PROGRAM main
  VAR
    B1 AT %IX0.0  : BOOL; (* sensor de piezas *)
    S1 AT %IX0.1  : BOOL; (* RESET *)
    KM1 AT %QX0.0 : BOOL; (* motor de la cinta *)
    H1 AT %QX0.1  : BOOL; (* caja llena *)
    PIEZAS        : CTU;
    LLENA         : BOOL;
    CUENTA        : INT; (* piezas en la caja *)
  END_VAR

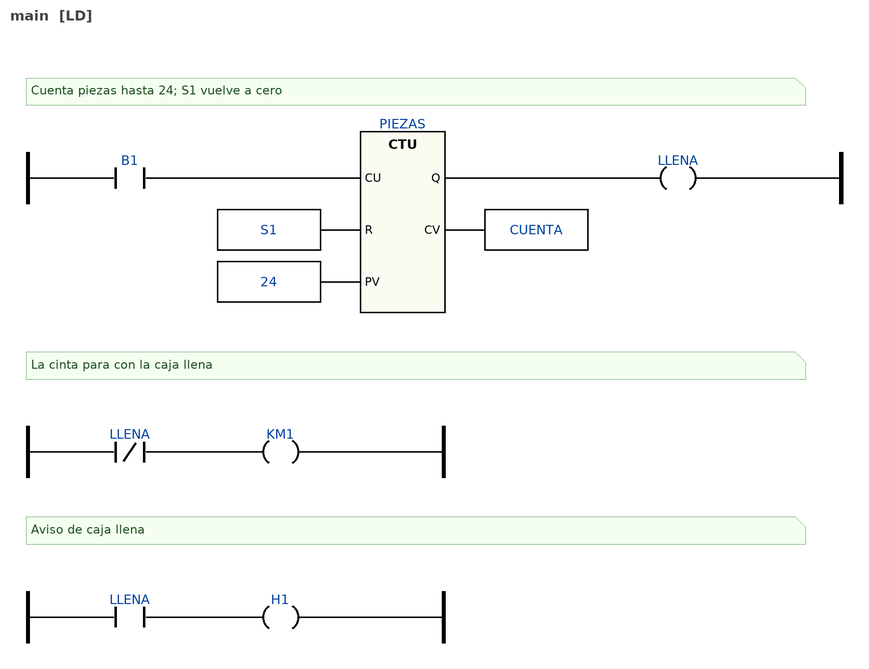
(* LD diagram, written out as Structured Text *)
(* Cuenta piezas hasta 24; S1 vuelve a cero *)
PIEZAS(CU := B1, R := S1, PV := 24);
LLENA := PIEZAS.Q;
CUENTA := PIEZAS.CV;
(* La cinta para con la caja llena *)
KM1 := NOT LLENA;
(* Aviso de caja llena *)
H1 := LLENA;
END_PROGRAM
